ABB RAPID module: BareProg1x.mod

%%%
  VERSION:1
  LANGUAGE:ENGLISH
%%%
MODULE MOD_BareProg1x

    ! -------------------------------
    ! Define customized variables here
    ! ...

	! Tool variables:

	! Reference variables:

	PROC Main()
		ConfJ \On;
		ConfL \Off;
		! Program generated by RoboDK v6.0.7 for ABB IRB 120-3/0.6 on XX/XX/XXXX 12:58:43
		! Using nominal kinematics.
		MoveAbsJ [[20.000000,-10.000000,20.000000,0.000000,30.000000,0.000000],[9E+09,9E+09,9E+09,9E+09,9E+09,9E+09]],v500,z1,tool0 \WObj:=wobj0;
		MoveAbsJ [[0.000000,-10.000000,20.000000,0.000000,30.000000,0.000000],[9E+09,9E+09,9E+09,9E+09,9E+09,9E+09]],v500,z1,tool0 \WObj:=wobj0;
	ENDPROC

ENDMODULE
